// TIA Portal V20 export
// export: Created 2026-10-19T18:02:23.5996088Z, ExportSetting WithDefaults, DisplayName Totally Integrated Automation Portal, DisplayVersion V20 Update 6, DisplayName TIA Portal Openness, DisplayVersion V20 Update 6, DisplayName TIA Portal Version Control Interface, DisplayVersion V20 Update 6, DisplayName SINAMICS Startdrive Advanced, DisplayVersion V20 SP1, DisplayName SINAMICS Startdrive G130, G150, S120, S150, SINAMICS MV, G220, S200, S210, DisplayVersion V20 SP1, DisplayName SINAMICS Startdrive G110M, G120, G120C, G120D, G120P, G115D, DisplayVersion V20 SP1, DisplayName STEP 7 Professional, DisplayVersion V20 Update 6, DisplayName STEP 7 Safety, DisplayVersion V20 Update 2, DisplayName WinCC Basic/Comfort/Advanced, DisplayVersion V20 Update 6, DisplayName WinCC Unified, DisplayVersion V20 Update 6
DATA_BLOCK "VTD_FB_DB"   // DB25
VERSION : 0.1
// stored: AutoNumber true, DBAccessibleFromOPCUA true, DBAccessibleFromWebserver true, InstanceOfName VTD_FB, InstanceOfType FB
"VTD_FB"
   // VAR_INPUT
   //    Cnv_Sensors : "ECnv_Inputs";
   //    VTD_Settings : "VTD_Settings";
   // END_VAR
   // VAR_IN_OUT
   //    VTD_Control : "VTD_Control";
   //    SinaSpeed : SinaSpeed;
   // END_VAR
   // VAR
   //    State : UInt;
   //    I_State : UInt;
   //    LD_Timer : TON_TIME;
   //    LP_Timer { S7_SetPoint := 'True'} : TON_TIME;
   //    Watchdog { S7_SetPoint := 'True'} : TON_TIME;
   //    CS_TImer { S7_SetPoint := 'True'} : TON_TIME;
   //    Interlock_Timer { S7_SetPoint := 'True'} : TON_TIME;
   //    MainSetpoint : Int;
   //    Position_Offset : Real;
   //    ChangeToLow : Array[1..4] of DInt;
   //    DestPosition : Real;
   //    SetUpSpeed : UInt;
   //    LevelBelowExtractor : UInt;
   //    IEC_Timer_0_Instance { S7_SetPoint := 'True'} : TON_TIME;
   //    DestinationLevel : UInt;
   //    CurrentlLevel : UInt;
   //    VTD_ID_Decoded { ExternalAccessible := 'False'; ExternalVisible := 'False'; ExternalWritable := 'False'} : "ID_Decoded";
   //    Cnv_ID_Decoded { ExternalAccessible := 'False'; ExternalVisible := 'False'; ExternalWritable := 'False'} : "ID_Decoded";
   //    IEC_Timer_0_Instance_1 { S7_SetPoint := 'True'} : TON_TIME;
   //    IEC_Timer_0_Instance_2 { S7_SetPoint := 'True'} : TON_TIME;
   //    VTD_ControlInstructionTask_ID_Old : Int;
   //    R_Execulte { S7_SetPoint := 'True'} : R_TRIG;
   // END_VAR
BEGIN
END_DATA_BLOCK
